(* IEC 61131-3 sources: yak/samples/x-iec-61131-3, 5 files *)

(* ---- ALMOnOff.st ---- *)
INTERFACE
    USES Define;
    FUNCTION_BLOCK MC_HandleALM;
END_INTERFACE

IMPLEMENTATION
// ============================================================================
// ----------- Function Blocks ------------------------------------------------
// ============================================================================

FUNCTION_BLOCK MC_HandleALM
// ----------------------------------------------------------------------------
//  <division / place / author>
// ----------------------------------------------------------------------------
//  Functionality description: This function block switches the active line
//                             module on/off. Also errors can be acknowledged.
// ----------------------------------------------------------------------------
//  Task assignment: This function block has to be used in cyclical tasks.
// ----------------------------------------------------------------------------
//  change log table:
//  version   date        expert in charge        changes applied
//  01.00.00  04.02.04    A. Krull A&D B18        created
//  02.00.00  08.11.04    S. Eisfeld A&D B18      alm not disabled when reset
//                                                occurs. With reset and enable
//                                                bit 1st error reset, 2nd
//                                                enable alm.
//  03.00.00  28.09.05    I. Hall SEA             Complete re-write to simplify operation

// ============================================================================
  VAR_INPUT
    ALMEnable    : BOOL; // rising edge 0->1: switch on active line module; falling edge: switch off
    PZDReceive   : WORD; // status word of active line module
  END_VAR

  VAR_OUTPUT

    PZDSend  : WORD; //command word of active line module
    ALMOn    : BOOL; //state of active line module (TRUE = On, FALSE = Off)
    ALMError : BOOL; //State of error (TRUE = error, FALSE = no error)

  END_VAR

  VAR
    ALMOnint    : BOOL; //state of active line module (TRUE = On, FALSE = Off)
    ALMErrorint : BOOL; //State of error (TRUE = error, FALSE = no error)
    retdint         :DINT ;

     END_VAR

//  get status of the ALM
   IF (PZDReceive AND 16#0017) = 16#0017 THEN
      ALMOn := TRUE;
      ALMOnint := TRUE;

  ELSE
      ALMOn := FALSE;
      ALMOnint := FALSE;
  END_IF;
  IF (PZDReceive AND 16#0008) = 16#0008 THEN
      ALMError := TRUE;
      ALMErrorint := TRUE;
  ELSE
      ALMError := FALSE;
      ALMErrorint := FALSE;
      //no error in status word -> reset acknowledge bit in command word
      PZDSend := PZDSend AND 16#FF7F;

  END_IF ;

 // Control of unit
    IF (ALMerrorint =  TRUE) AND (ALMENABLE  = TRUE) THEN
      PZDSend := PZDSend OR 16#0080; //reset error

      RetDINT := _waittime(T#50ms); // wait
      PZDSend := PZDSend OR 16#040A ;//AND 16#FFFE; // send disable command
      RetDINT := _waittime(T#100ms); // wait
      PZDSend := PZDSend OR 16#040b; // send enable command (see a rising edge)
     // stateNumber := 0;
END_IF ;
    IF ALMEnable = FALSE THEN
      PZDSend := PZDSend AND 16#FFFE; //disable ALM

  END_IF ;

     IF (ALMEnable = TRUE)  AND (PZDReceive = 16#0250)  THEN
      PZDSend := 16#040A ; //give ALM an off command so as to be able to give it a rising edge start command
      RetDINT := _waittime(T#200ms); // wait
  END_IF ;

      IF (PZDRECEIVE = 16#211)  THEN //wait for acknowledge of previous command
      RetDINT := _waittime(T#50ms); // wait
      PZDSend := PZDSend OR 16#040b ; // start alm
END_IF ;

END_FUNCTION_BLOCK

END_IMPLEMENTATION

(* ---- motorek.plc ---- *)
FUNCTION shr: BYTE
	VAR_INPUT
		in: BYTE;
		nr: BYTE;
	END_VAR

loop:
	LD	nr
	EQ	0
	RETC

	LD	nr
	SUB	1
	ST	nr

	LD	in
	DIV	2
	ST	in
	ST	shr

	JMP	loop
END_FUNCTION

FUNCTION_BLOCK pwm
	VAR_INPUT
		pwmval: INT;
	END_VAR
	VAR_EXTERNAL
		Forward: BOOL;
		Backward: BOOL;
	END_VAR
	VAR
		cc: INT := 0;
		runback: BOOL;
	END_VAR

	LD	pwmval
	LT	0
	ST	runback

	JMPCN	runpwm

	LD	pwmval
	STN	pwmval

runpwm:
	LD	pwmval
	GE	100
	JMPCN	cont

	LD	99
	ST	pwmval
cont:
	LD	cc
	ADD	1
	ST	cc

	EQ	100
	JMPCN	norst

	LD	0
	ST	cc

norst:	LD	cc
	GE	pwmval

	JMPC	pwm2

	LD	runback

	JMPCN	fwd

	S	Backward
	R	Forward

	RETC

fwd:
	LD	1
	S	Forward
	R	Backward

	RET

pwm2:	LD	1
	R	Forward
	R	Backward

	RET

END_FUNCTION_BLOCK

PROGRAM prg_motorek
	VAR
		controler: PID;
		dopwm:	pwm;
		spwm: INT := 0;
	END_VAR
	VAR_EXTERNAL
		P: DINT;
		I: DINT;
		D: DINT;

		ISAT: DINT;

		Forward: BOOL;
		SP: DINT;

		RPS: DINT;
	END_VAR

	LD	P
	ST	controler.P
	LD	I
	ST	controler.I
	LD	D
	ST	controler.D
	LD	ISAT
	ST	controler.ISAT

	LD	SP
	SUB	RPS

	ST	controler.PV

	CAL	controler

	LD	controler.AV
	ST	spwm

exepwm:
	CAL	dopwm(PWMVal := spwm)
END_PROGRAM

(* Program for measurement of rotations per sec *)
(* Forward:  00 10 11 01 00 *)
(* Backward: 00 01 11 10 00 *)
PROGRAM prg_otacky
	VAR
		CONSTANT StateMask: BYTE := 16#30;
		StateOld: BYTE := 0;
		StateNew: BYTE;
		TimeOld: DINT := 0;
		Otacky: DINT := 0;
		citac: DINT := 0;
	END_VAR

	VAR_EXTERNAL
		Direction: BOOL;
		StateInput: BYTE;
		time: DINT;
		RPS: DINT;
	END_VAR

	LD	StateInput
	AND	StateMask

	shr	4

	ST	StateNew
	EQ	StateOld
	RETC

	LD	StateNew
	EQ	0
	JMPCN	Test2

	LD	StateOld
	EQ	1
	ST	Direction

	JMP	SaveState

Test2:	LD	StateNew
	EQ	2
	JMPCN	Test3

	LD	StateOld
	EQ	0
	ST	Direction

	JMP	SaveState

Test3:	LD	StateNew
	EQ	3
	JMPCN	Test4

	LD	StateOld
	EQ	2
	ST	Direction

	JMP	SaveState

Test4:	LD	StateNew
	EQ	1
	JMPCN	SaveState

	LD	StateOld
	EQ	3
	ST	Direction

SaveState:
	LD	StateNew
	ST	StateOld

	LD	citac
	ADD	1
	ST	citac

	EQ	4
	RETCN

	LD	0
	ST	citac

	LD	time
	SUB	TimeOld
	MUL	4

	ST	Otacky
	EQ	0
	RETC

	LD	10000
	DIV	Otacky
	ST	RPS

	LD	time
	ST	TimeOld

	LD	Direction
	RETC

	LD	RPS
	STN	RPS
END_PROGRAM

PROGRAM	prg_time
	VAR_EXTERNAL
		time: DINT;
	END_VAR

	LD	time
	ADD	1
	ST	time
END_PROGRAM

CONFIGURATION motorek
	VAR_GLOBAL
		time: DINT := 0;
		RPS AT %QB10: DINT := 0;

		SP AT %IB10: DINT;

		(* *)
		Forward AT %Q0.0: BOOL := FALSE;
		Backward AT %Q0.1: BOOL := FALSE;

		StateInput AT %IB0: BYTE;

		(* TRUE - otaceni vpred, FALSE - otaceni vzad *)
		Direction: BOOL := FALSE;

		(* Constants for PID controler *)
		P: DINT := 4;
		I: DINT := 1;
		D: DINT := 2;

		ISAT: DINT := 100;
	END_VAR

	RESOURCE xx ON yy
		TASK rustTask(INTERVAL:=T#10ms);
		TASK measureRotationTask(SINGLE:=%I1.0);
		TASK measureRPSTask(INTERVAL:=T#0.1ms);

		PROGRAM p1 WITH rustTask: prg_motorek();
		PROGRAM p2 WITH measureRotationTask: prg_otacky();
		PROGRAM p3 WITH measureRPSTask: prg_time();
	END_RESOURCE
END_CONFIGURATION

(* ---- PKG41.st ---- *)
INTERFACE

    USEPACKAGE cam;

    // USES header;

    // USELIB testlib;

    VAR_GLOBAL CONSTANT
           PI : REAL := 3.1415;
           ARRAY_MAX : INT := 3;
    END_VAR

    TYPE
        array1dim : ARRAY [0..ARRAY_MAX] OF INT;
        array2dim : ARRAY [0..3] OF array1dim;
        enumTrafficLight : (RED, YELLOW, GREEN);

        structCollection : STRUCT
            toAxisX : posaxis;
            aInStruct1dim : array1dim;
            eTrafficInStruct : enumTrafficLight;
            iCounter : INT;
            bStatus : WORD;
        END_STRUCT;

        arrayOfStruct : ARRAY [0..5] OF structCollection;

    END_TYPE

    // *****************************************************
    // * Variablendeklaration im INTERFACE                 *
    // *****************************************************)

    VAR_GLOBAL

        g_aMyArray : ARRAY [0..11] OF REAL := [3 (2(4), 2(18))];

        g_aMy2dim : array2dim;

        g_aMy1dim : array1dim;

        g_sMyStruct : structCollection;

        g_aMyArrayOfStruct : arrayOfStruct;

        g_tMyTime : TIME := T#0d_1h_5m_17s_4ms;

        g_eMyTraffic : enumTrafficLight := RED;

        g_iMyInt : INT := -17;
    END_VAR

    VAR_GLOBAL RETAIN
    END_VAR

    FUNCTION_BLOCK FB_myFirst;
    FUNCTION FC_myFirst;
    PROGRAM myPRG;

END_INTERFACE

// *****************************************************
// * IMPLEMENTATION-Teil                               *
// *****************************************************

IMPLEMENTATION

    VAR_GLOBAL CONSTANT
    END_VAR

    TYPE
    END_TYPE

    VAR_GLOBAL
        g_boDigInput1 : BOOL;
    END_VAR

    VAR_GLOBAL RETAIN
    END_VAR

    EXPRESSION xCond
        xCond := g_boDigInput1;
    END_EXPRESSION

    // *****************************************************
    // * FUNCTION_BLOCK                                    *
    // *****************************************************)

    FUNCTION_BLOCK FB_myFirst

        VAR CONSTANT
        END_VAR

        TYPE
        END_TYPE

        VAR_INPUT
        END_VAR

        VAR_IN_OUT
        END_VAR

        VAR_OUTPUT
        END_VAR

        VAR
        END_VAR

        VAR_TEMP
        END_VAR

        g_eMyTraffic := GREEN; // z.B. Umschalten der Ampel

    END_FUNCTION_BLOCK

    // *****************************************************
    // * FUNCTION                                          *
    // *****************************************************)

    FUNCTION FC_myFirst : INT

        VAR CONSTANT
        END_VAR

        TYPE
        END_TYPE

        VAR_INPUT
        END_VAR

        VAR
        END_VAR

        g_eMyTraffic := YELLOW;

        FC_myFirst := 17;

    END_FUNCTION

    // *****************************************************
    // * PROGRAM                                           *
    // *****************************************************

    PROGRAM myPRG

        VAR CONSTANT
        END_VAR

        TYPE
        END_TYPE

        VAR
            instFBMyFirst : FB_myFirst;

            retFCMyFirst : INT;
        END_VAR

        VAR_TEMP
        END_VAR

        instFBMyFirst ();

        retFCMyFirst := FC_myFirst ();

        WAITFORCONDITION xCond WITH TRUE DO
            ;
        END_WAITFORCONDITION;

    END_PROGRAM

END_IMPLEMENTATION

(* ---- snake.plc ---- *)
FUNCTION shl:BYTE
	VAR_INPUT
		in: BYTE;
	END_VAR

	LD	in
	MUL	2
	ST	shl
END_FUNCTION

FUNCTION_BLOCK rust
	VAR_INPUT
		in: BYTE;
	END_VAR
	VAR_OUTPUT
		out: BYTE;
	END_VAR
	VAR
		mask: BYTE := 1;
	END_VAR

	LD	in
	OR	mask
	ST	out

	LD	mask
	MUL	2
	ST	mask

	LD	mask
	EQ	0

	RETCN

	LD	1
	ST	mask
END_FUNCTION_BLOCK

PROGRAM prg_rust
	VAR_IN_OUT
		outx: BYTE;
	END_VAR
	VAR
		r: rust;
	END_VAR
	VAR_EXTERNAL
		out: BYTE;
		rust: BOOL;
		rotace: BOOL;
	END_VAR

	LD	outx
	EQ	16#ff
	JMPCN	volej
	LD	0
	ST	outx

	(* switch to second effect *)
	R	rust
	S	rotace

volej:	LD	outx
	ST	r.in
	CAL	r
	LD	r.out
	ST	outx
	RET

END_PROGRAM

PROGRAM prg_light1
	VAR_EXTERNAL
		out: BYTE;
	END_VAR

	LD	2#10101010
	ST	out
END_PROGRAM

PROGRAM prg_light2
	VAR_EXTERNAL
		out: BYTE;
	END_VAR

	LD	2#01010101
	ST	out
END_PROGRAM

PROGRAM prg_rotace
	VAR_EXTERNAL
		out: BYTE;
		rust: BOOL;
		rotace: BOOL;
	END_VAR

	LD	out
	shl
	ST	out
	EQ	0
	RETCN
	LD	1
	ST	out

	(* Switch to second effect *)
	R	rotace
	S	rust
END_PROGRAM

CONFIGURATION snake
	VAR_GLOBAL
		out AT %QB0: BYTE := 1;
		rust: BOOL := FALSE;
		rotace AT %MX0.0: BOOL := TRUE;
	END_VAR

	RESOURCE xx ON yy
		TASK rustTask(SINGLE := rust, INTERVAL:=T#0.5s);
		TASK rotaceTask(SINGLE := %MX0.0, INTERVAL:=T#0.5s);
		TASK ligthTask(SINGLE := rotace);
		TASK ligthTask2(SINGLE := rust);

		PROGRAM p1 WITH rustTask: prg_rust(outx:=out);
		PROGRAM p2 WITH rotaceTask: prg_rotace();
(*		PROGRAM p3 WITH ligthTask: prg_light1(); *)
(*		PROGRAM p4 WITH ligthTask2: prg_light2(); *)
	END_RESOURCE
END_CONFIGURATION

(* ---- chaser_st.st ---- *)
FUNCTION SCROLL_LEFT: INT
  (* Interface *)
  VAR_IN_OUT
    bits: INT;
  END_VAR  (* Local Vars. *)
  VAR_INPUT
    top_bit: INT;
  END_VAR

  bits := bits * 2;

  IF (bits >= top_bit)
  THEN
    bits := bits + 1 - top_bit;
  END_IF;

  SCROLL_LEFT := bits;
END_FUNCTION

FUNCTION SCROLL_RIGHT: INT
  VAR_IN_OUT
    bits: INT;
  END_VAR
  VAR_INPUT
    top_bit: INT;
  END_VAR

  IF ((bits mod 2) = 0)
    THEN top_bit := 0;
  END_IF;

  bits := bits / 2;
  bits := bits + top_bit/2;

  SCROLL_RIGHT := bits;

END_FUNCTION

PROGRAM SCROLL
  VAR_EXTERNAL
    left_bt  : BOOL;
    right_bt : BOOL;
    bits : INT;
  END_VAR
  VAR
    (* We don't suport passing external type variables to functions *)
    (* I (Mario) don't have time to fix this
     * and would like to commit something before I do go on holidays.
     * So for now, we use this workaround...
     *)
    local_bits : INT;
    direction : BOOL; (* FALSE is right, TRUE is left , we do not yet support enums *)
  END_VAR

  IF left_bt  THEN direction := FALSE; END_IF;
  IF right_bt THEN direction := TRUE;  END_IF;

  local_bits := bits;
  IF direction
    THEN bits := SCROLL_LEFT(local_bits, 16);
    ELSE bits := SCROLL_RIGHT(local_bits, 16);
  END_IF;

END_PROGRAM

CONFIGURATION config1
  VAR_GLOBAL
    bits AT %L : INT := 1;
    left_bt  AT %left  : BOOL;
    right_bt AT %right : BOOL;
   END_VAR

  PROGRAM main: SCROLL(left_bt := left_bt, right_bt := right_bt, bits := bits);
END_CONFIGURATION
